ACTION LastComp_active:
wButtonColor:=16#FF00FFFF;

sStateDescription	:=	'Finish';
sStateInstructions	:= 	'LastComponentMixed';

bDisableAmount	:=FALSE;
bDisableName	:=FALSE;
bDisableTime	:=FALSE;
END_ACTION

ACTION LastComp_exit:
VisuElems.CurrentVisu:= 'StartVisu';
stTriblender.bDisolvingDone:=TRUE;
END_ACTION

ACTION MixComponent_active:
sStateDescription	:=	'Component Inside';
sStateInstructions	:= 	'Insert component in
 the specified amount';
END_ACTION

ACTION MixComponent_entry:
bContinue:=FALSE;

bDisableAmount	:=FALSE;
bDisableName	:=FALSE;
bDisableTime	:=FALSE;

wButtonColor:=16#FFFF0000;
IF iCurrentMixingComponent<g_Prod.cMaxCompInProduct-1 THEN
	stTriblender.bLastComponent:=NOT arrComponents[iCurrentMixingComponent+1].bComponentEnable;
END_IF
stTriblender.sComponenetAmount:=TO_STRING(arrComponents[iCurrentMixingComponent].rCompActWeight);
stTriblender.sComponenetName:=arrComponents[iCurrentMixingComponent].sDescription;
stTriblender.tComponenetMixingTime:=TO_TIME(arrComponents[iCurrentMixingComponent].iMixingTime*1000);
fb_TriBlenderPump.m_Run(RPM:=arrComponents[iCurrentMixingComponent].rRpmTarget);
END_ACTION

ACTION MixDoneWaitAnother_active:
sStateDescription	:='Triblender valve Opened';
sStateInstructions	:= 'Mix Component done,
 open triblender valve';
END_ACTION

ACTION MixDoneWaitAnother_entry:
bContinue:=FALSE;

bDisableAmount:=TRUE;
bDisableName:=TRUE;
bDisableTime:=TRUE;
bDisableButton:=FALSE;
VisuElems.CurrentVisu:= 'StartVisu';



wButtonColor:=16#FF00FF00;
END_ACTION

ACTION OpenValve_entry:
bContinue:=FALSE;

bDisableAmount:=TRUE;
bDisableName:=TRUE;
bDisableTime:=TRUE;
bDisableButton:=FALSE;

tonStageCirculation(IN:=FALSE);


sStateDescription	:='Triblender valve Opened';
sStateInstructions	:= 'Open triblender valve';

wButtonColor:=16#FF00FF00;
END_ACTION

TRANSITION trans_RpmInTarget:
fb_TriBlenderPump.nRPM< arrComponents[i].rRpmTarget+10 and fb_TriBlenderPump.nRPM> arrComponents[i].rRpmTarget-10
END_TRANSITION

TRANSITION transCircDone:
tonStageCirculation.Q and stTriblender.rMaxAllowedPressure> stTriblender.rPressure and stTriblender.rMinAllowedFlow< stTriblender.rFlow
END_TRANSITION

ACTION WaitForDone_active:
tonStageCirculation(IN:= TRUE,PT:=stTriblender.tComponenetMixingTime);
iCirculationTimeLeft:= TO_UINT(tonStageCirculation.PT - tonStageCirculation.ET)/1000;
bDisableButton:=TRUE;
END_ACTION

ACTION WaitForDone_entry:
wButtonColor:=16#FF0000FF;

sStateDescription	:=	'Waiting';
sStateInstructions	:= 	'Wait for mixing done';
bContinue:=FALSE;

bDisableAmount	:=FALSE;
bDisableName	:=FALSE;
bDisableTime	:=FALSE;


tonStageCirculation(IN:= FALSE);
END_ACTION

ACTION WaitForDone_exit:
stTriblender.bComponenetMixDone:=TRUE;
wButtonColor:=16#FF00FF00;

bDisableAmount	:=TRUE;
bDisableName	:=TRUE;
bDisableTime	:=TRUE;


tonStageCirculation(IN:= FALSE);
END_ACTION

ACTION WaitForStartPump_active:
sStateDescription	:='Start Water Circulation';
sStateInstructions	:= 'Start water circulation, check for leaks';
iCurrentMixingComponent:=0;
bContinue:=FALSE;
FOR i:= 0 TO g_Prod.cMaxCompInProduct-1 DO
	IF arrComponents[i].bIsWater THEN
		fb_TriBlenderPump.m_Run(RPM:=arrComponents[i].rRpmTarget);
	END_IF
END_FOR

wButtonColor:=16#FFFF0000;
END_ACTION

ACTION WaitForStartPump_entry:

stTriblender.bStartDisolving:=FALSE;
END_ACTION

ACTION WaterCirculation_active:
tonStageCirculation(IN:= stTriblender.bPumpOnFdbk,PT:=stTriblender.tWaterCirculationTimeout);
iCirculationTimeLeft:= TO_UINT(tonStageCirculation.PT - tonStageCirculation.ET)/1000;

bDisableButton:=TRUE;

sStateDescription	:='Wait for pressure and flow';
sStateInstructions	:= 'Water circulation in progress,
 check for leaks';
END_ACTION

ACTION WaterCirculation_entry:
bContinue:=FALSE;


bDisableAmount:=TRUE;
bDisableName:=TRUE;
bDisableTime:=FALSE;

tonStageCirculation(IN:=FALSE);
END_ACTION

ACTION WaterCirculation_exit:
tonStageCirculation(IN:=FALSE);
END_ACTION

END_PROGRAM

// ---- 03 Project/23 CIP/FB_Fill_Water.TcPOU
FUNCTION_BLOCK FB_Fill_Water EXTENDS FB_SFC_Cycle
VAR_INPUT
	valve : E_Pis_Name;;
	reqLevel: REAL;
	actLevel: REAL;
	
	fillCondition: BOOL;


END_VAR
VAR_OUTPUT
END_VAR
VAR
	fbHysteresis: FB_Hysteresis_REAL;
	stValve: REFERENCE TO ST_Piston;

END_VAR

stValve REF= stPis[valve];
IF NOT __ISVALIDREF(stValve) THEN;
	RETURN;
END_IF

fbHysteresis(
	fIn:= , 
	fHigh:= reqLevel, 
	fLow:= reqLevel-50.0, 
	iDigitsAfterDot:= , 
	bOut=> );

IF stValve.st_Open 
AND (NOT fbHysteresis.bOut
OR NOT fillCondition)
THEN;
	stValve.req_Close:=TRUE;
	
ELSIF stValve.st_Close 
AND fbHysteresis.bOut
THEN;
	stValve.req_Open:=TRUE;
END_IF

END_FUNCTION_BLOCK

// ---- 00 Library/01 Piston/TextList_Piston_Recipe_State.TcTLO
TEXTLIST TextList_Piston_Recipe_State
  0 = ' '
  1 = 'Open'
  2 = 'Close'
   = ''
END_TEXTLIST

// ---- 00 Library/01 Piston/TextList_Piston_Recipe_State_CloseOpen.TcTLO
TEXTLIST TextList_Piston_Recipe_State_CloseOpen
  0 = ' '
  1 = 'Close'
  2 = 'Open'
   = ''
END_TEXTLIST

// ---- 00 Library/01 Piston/TextList_Piston_Recipe_State_DownUp.TcTLO
TEXTLIST TextList_Piston_Recipe_State_DownUp
  0 = ' '
  1 = 'Down'
  2 = 'Up'
   = ''
END_TEXTLIST

// ---- 00 Library/01 Piston/TextList_Piston_Recipe_State_InOut.TcTLO
TEXTLIST TextList_Piston_Recipe_State_InOut
  0 = ' '
  1 = 'In'
  2 = 'Out'
   = ''
END_TEXTLIST

// ---- 00 Library/01 Piston/TextList_Piston_Recipe_State_OnOff.TcTLO
TEXTLIST TextList_Piston_Recipe_State_OnOff
  0 = ' '
  1 = 'On'
  2 = 'Off'
   = ''
END_TEXTLIST

// ---- 00 Library/01 Piston/TextList_Piston_Recipe_State_OpenClose.TcTLO
TEXTLIST TextList_Piston_Recipe_State_OpenClose
  0 = ' '
  1 = 'Open'
  2 = 'Close'
   = ''
END_TEXTLIST

// ---- 00 Library/01 Piston/TextList_Piston_Recipe_State_UpDown.TcTLO
TEXTLIST TextList_Piston_Recipe_State_UpDown
  0 = ' '
  1 = 'Up'
  2 = 'Down'
   = ''
END_TEXTLIST

// ---- 00 Library/01 Piston/VISU/vis_Piston_Control1.TcVIS
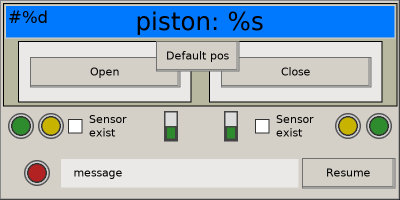
VISUALIZATION vis_Piston_Control1  // 400x200
VAR_IN_OUT
	stPis: ST_Piston;
END_VAR
    Rectangle (0,0 400x200)
    Rectangle (3,3 394x103), colour toggle: NOT stPis.b_Enable
    Rectangle (18,41 173x61), colour toggle: stPis.st_Open
    Rectangle (209,41 173x61), colour toggle: stPis.st_Close
    Button (30,57 150x30), "Open", colour toggle: stPis.req_Open, input disabled if: stPis.b_DeactivateMan OR NOT stPis.b_InterLock_Open
        toggle stPis.req_OpenMan
    Button (221,57 150x30), "Close", colour toggle: stPis.req_Close, input disabled if: stPis.b_DeactivateMan OR NOT stPis.b_InterLock_Close
        toggle stPis.req_CloseMan
    DipSwitch (156,111 30x30), tooltip "Open Sensor state", variable: stPis.sen_Open, invisible if: NOT stPis.sen_Open_Exist, behaviour: TOGGLE, style: Switch-DipSwitch-Green
    DipSwitch (216,111 30x30), tooltip "Close Sensor state", variable: stPis.sen_Close, invisible if: NOT stPis.sen_Close_Exist, behaviour: TOGGLE, style: Switch-DipSwitch-Green
    Checkbox (66,108 99x36), "Sensor exist", variable: stPis.sen_Open_Exist
    Checkbox (253,108 99x36), "Sensor exist", variable: stPis.sen_Close_Exist
    Lamp1 (6,111 30x30), tooltip "Open sensor", variable: stPis.sen_Open, invisible if: NOT stPis.sen_Open_Exist, style: Lamp-Lamp1-Green
    Lamp1 (333,111 30x30), tooltip "Close valve", variable: stPis.valve_Close, style: Lamp-Lamp1-Yellow
    Lamp1 (22,158 30x30), tooltip "Error", variable: stPis.b_Error, style: Lamp-Lamp1-Red
    Textfield (60,158 239x30), "message"
    Button (302,158 93x30), "Resume", colour toggle: stPis.b_Error
        toggle stPis.b_Resume
    Button (156,41 83x30), "Default pos", colour toggle: stPis.req_DefaultPos, input disabled if: stPis.b_DeactivateMan
        toggle stPis.req_DefaultPos
    Textfield (5,5 390x33), "piston: %s", text variable: stPis.sName
    Textfield (5,7 42x21), "#%d", text variable: stPis.iPisNum
    Lamp1 (36,111 30x30), tooltip "Open valve", variable: stPis.valve_Open, style: Lamp-Lamp1-Yellow
    Lamp1 (364,111 30x30), tooltip "Close sensor", variable: stPis.sen_Close, invisible if: NOT stPis.sen_Close_Exist, style: Lamp-Lamp1-Green
END_VISUALIZATION

// ---- 00 Library/01 Piston/VISU/vis_Piston_Control1_Compact.TcVIS
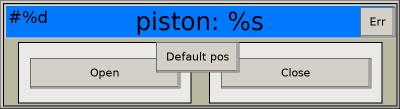
VISUALIZATION vis_Piston_Control1_Compact  // 400x109
VAR_IN_OUT
	stPis: ST_Piston;
END_VAR
    Rectangle (0,0 400x109)
    Rectangle (3,3 394x103), colour toggle: NOT stPis.b_Enable
    Rectangle (18,42 173x61), colour toggle: stPis.st_Open
    Rectangle (209,42 173x61), colour toggle: stPis.st_Close
    Button (30,58 150x30), "Open", colour toggle: stPis.req_Open, input disabled if: stPis.b_DeactivateMan OR NOT stPis.b_InterLock_Open
        toggle stPis.req_OpenMan
    Button (221,58 150x30), "Close", colour toggle: stPis.req_Close, input disabled if: stPis.b_DeactivateMan OR NOT stPis.b_InterLock_Close
        toggle stPis.req_CloseMan
    Button (156,42 83x30), "Default pos", colour toggle: stPis.req_DefaultPos, input disabled if: stPis.b_DeactivateMan
        toggle stPis.req_DefaultPos
    Textfield (5,5 390x33), "piston: %s", text variable: stPis.sName
    Textfield (5,7 42x21), "#%d", text variable: stPis.iPisNum
    Button (360,7 35x30), "Err", colour toggle: stPis.b_Error
        toggle stPis.b_Resume
END_VISUALIZATION

// ---- 00 Library/01 Piston/VISU/vis_Piston_Control2_CloseOpen.TcVIS
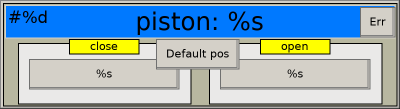
VISUALIZATION vis_Piston_Control2_CloseOpen  // 400x109
VAR_IN_OUT
	stPis			: ST_Piston;
END_VAR
VAR_INPUT
	sLable_Open		: STRING:='lable open';
	sLable_Close	: STRING:='lable close';
END_VAR
    Rectangle (0,0 400x109)
    Rectangle (3,3 394x103), colour toggle: NOT stPis.b_Enable
    Rectangle (209,43 173x61), colour toggle: stPis.st_Open
    Button (220,59 150x30), "%s", text variable: sLable_Open, colour toggle: stPis.req_Open, input disabled if: stPis.b_DeactivateMan OR NOT stPis.b_InterLock_Open
        toggle stPis.req_OpenMan
    RoundedRectangle (260,39 70x15), "open"
    Rectangle (18,43 173x61), colour toggle: stPis.st_Close
    Button (29,59 150x30), "%s", text variable: sLable_Close, colour toggle: stPis.req_Close, input disabled if: stPis.b_DeactivateMan OR NOT stPis.b_InterLock_Close
        toggle stPis.req_CloseMan
    RoundedRectangle (69,39 70x15), "close"
    Button (156,39 83x30), "Default pos", colour toggle: stPis.req_DefaultPos, input disabled if: stPis.b_DeactivateMan
        toggle stPis.req_DefaultPos
    Textfield (5,5 390x33), "piston: %s", text variable: stPis.description
    Textfield (5,7 42x21), "#%d", text variable: stPis.iPisNum
    Button (360,7 35x30), "Err", colour toggle: stPis.b_Error
        toggle stPis.b_Resume
END_VISUALIZATION

// ---- 00 Library/01 Piston/VISU/vis_Piston_Control2_OpenClose.TcVIS
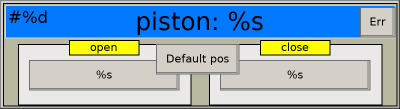
VISUALIZATION vis_Piston_Control2_OpenClose  // 400x109
VAR_IN_OUT
	stPis			: ST_Piston;
END_VAR
VAR_INPUT
	sLable_Open		: STRING:='lable open';
	sLable_Close	: STRING:='lable close';
END_VAR
    Rectangle (0,0 400x109)
    Rectangle (3,3 394x103), colour toggle: NOT stPis.b_Enable
    Rectangle (18,44 173x61), colour toggle: stPis.st_Open
    Rectangle (209,44 173x61), colour toggle: stPis.st_Close
    Button (29,60 150x30), "%s", text variable: sLable_Open, colour toggle: stPis.req_Open, input disabled if: stPis.b_DeactivateMan OR NOT stPis.b_InterLock_Open
        toggle stPis.req_OpenMan
    Button (220,60 150x30), "%s", text variable: sLable_Close, colour toggle: stPis.req_Close, input disabled if: stPis.b_DeactivateMan OR NOT stPis.b_InterLock_Close
        toggle stPis.req_CloseMan
    Button (156,44 83x30), "Default pos", colour toggle: stPis.req_DefaultPos, input disabled if: stPis.b_DeactivateMan
        toggle stPis.req_DefaultPos
    RoundedRectangle (69,40 70x15), "open"
    RoundedRectangle (260,40 70x15), "close"
    Textfield (5,5 390x33), "piston: %s", text variable: stPis.description
    Textfield (5,7 42x21), "#%d", text variable: stPis.iPisNum
    Button (360,7 35x30), "Err", colour toggle: stPis.b_Error
        toggle stPis.b_Resume
END_VISUALIZATION

// ---- 00 Library/01 Piston/VISU/vis_Piston_Select.TcVIS
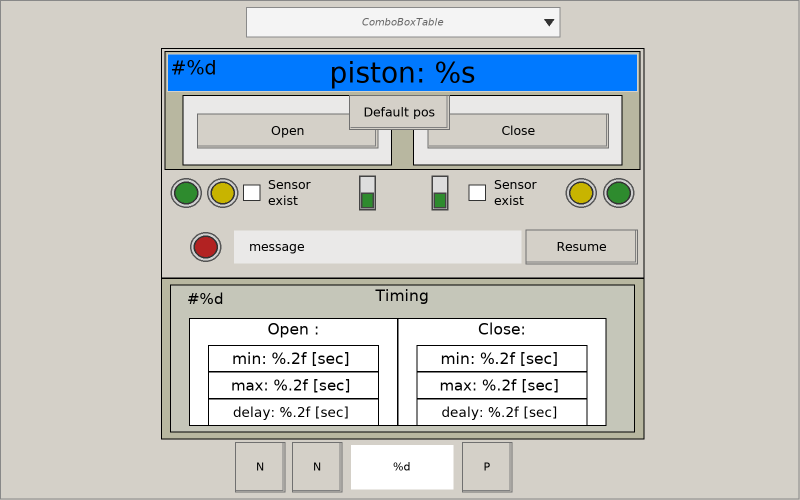
VISUALIZATION vis_Piston_Select  // 800x500
    Frame (161,48 483x230)
        shows vis_Piston_Control1(stPis := stPis[iPis_sel])
    Frame (161,278 483x161)
        shows vis_Piston_Times(stPis := stPis[iPis_sel])
    Button (292,442 50x50), "N"
        tap prg_Piston.bPis_Next_N
    Button (462,442 50x50), "P"
        tap prg_Piston.bPis_Next_P
    Textfield (350,444 104x46), "%d", text variable: iPis_sel
    ComboBoxTable (246,7 314x30), variable: iPis_sel, data array: g_Piston.arPisName
        p3854506369: g_Piston.arPisName[INDEX].Num
        p1892666644: g_Piston.arPisName[INDEX].Description
    Button (235,442 50x50), "N"
        tap prg_Piston.bPis_Next_N
END_VISUALIZATION

// ---- 00 Library/01 Piston/VISU/vis_Piston_Select_1.TcVIS
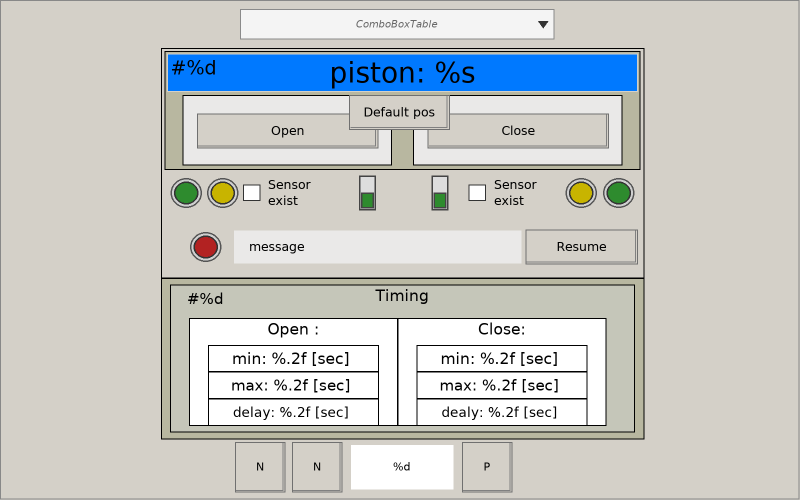
VISUALIZATION vis_Piston_Select_1  // 800x500
    Frame (161,48 483x230)
        shows vis_Piston_Control1(stPis := stPis[iPis_sel])
    Frame (161,278 483x161)
        shows vis_Piston_Times(stPis := stPis[iPis_sel])
    Button (292,442 50x50), "N"
        tap prg_Piston.bPis_Next_N
    Button (462,442 50x50), "P"
        tap prg_Piston.bPis_Next_P
    Textfield (350,444 104x46), "%d", text variable: iPis_sel
    ComboBoxTable (240,9 314x30), variable: iPis_sel, data array: arPisName
        p1128707560: C_MAX_Pistons_Exist
        p3854506369: arPisName[INDEX].Num
        p1892666644: arPisName[INDEX].Description
    Button (235,442 50x50), "N"
        tap prg_Piston.bPis_Next_N
END_VISUALIZATION

// ---- 00 Library/01 Piston/VISU/vis_Piston_Setting_Table.TcVIS
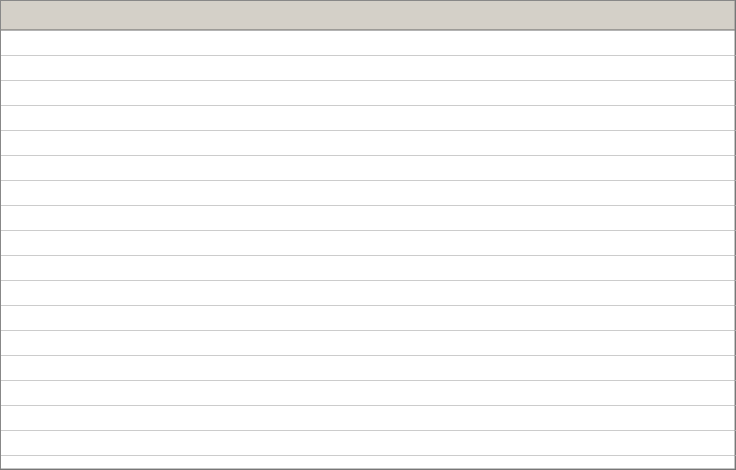
VISUALIZATION vis_Piston_Setting_Table  // 736x470
    Table (0,0 736x470), data array: stPisSetting
        p3854506369: stPisSetting[INDEX].t_minOpen
        p1892666644: stPisSetting[INDEX].t_minClose
        p338671338: stPisSetting[INDEX].t_maxOpen
        p2170511999: stPisSetting[INDEX].t_maxClose
        p3723444502: stPisSetting[INDEX].t_DelayOpen
        p1218418051: stPisSetting[INDEX].t_DelayClose
        p746581629: stPisSetting[INDEX].sen_Open_Exist
        p3104783080: stPisSetting[INDEX].sen_Close_Exist
END_VISUALIZATION

// ---- 00 Library/01 Piston/VISU/vis_Piston_Times.TcVIS
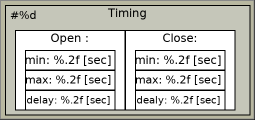
VISUALIZATION vis_Piston_Times  // 255x120
VAR_IN_OUT
	stPis: ST_Piston;
END_VAR
    Rectangle (0,0 255x120)
    Rectangle (5,5 245x110), "Timing"
    Rectangle (15,30 110x80), "Open :"
    Rectangle (125,30 110x80), "Close:"
    Rectangle (135,50 90x20), "min: %.2f [sec]", text variable: stPis.t_minClose
        OnMouseDown: write the text variable via Edit, min 0
    Rectangle (135,70 90x20), "max: %.2f [sec]", text variable: stPis.t_maxClose
        OnMouseDown: write the text variable via Edit, min 0
    Rectangle (25,70 90x20), "max: %.2f [sec]", text variable: stPis.t_maxOpen
        OnMouseDown: write the text variable via Edit, min 0
    Rectangle (25,50 90x20), "min: %.2f [sec]", text variable: stPis.t_minOpen
        OnMouseDown: write the text variable via Edit, min 0
    Rectangle (25,90 90x20), "delay: %.2f [sec]", text variable: stPis.t_DelayOpen
        OnMouseDown: write the text variable via Edit, min 0
    Rectangle (135,90 90x20), "dealy: %.2f [sec]", text variable: stPis.t_DelayClose
        OnMouseDown: write the text variable via Edit, min 0
    Textfield (4,5 39x21), "#%d", text variable: stPis.iPisNum
END_VISUALIZATION

// ---- 00 Library/03 SFC/vis_Cycle_Control.TcVIS
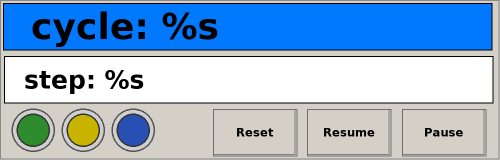
VISUALIZATION vis_Cycle_Control  // 500x160
VAR_IN_OUT
	fb: FB_SFC_Cycle;
END_VAR
VAR_INPUT
	sName: STRING:='Cycle name';
END_VAR
    Lamp1 (8,105 50x50), tooltip "Ready", variable: fb.bReady, style: Lamp-Lamp1-Green
    Lamp1 (108,105 50x50), tooltip "Done", variable: fb.bDone, style: Lamp-Lamp1-Blue
    Lamp1 (58,105 50x50), tooltip "Run", variable: fb.bRun, style: Lamp-Lamp1-Yellow
    RoundedRectangle (3,3 489x47), "cycle: %s", tooltip "POU name: %s", text variable: sName
        p4168582468: fb.refSFC.SFCErrorPOU
    RoundedRectangle (4,56 489x47), "step: %s", text variable: fb.refSFC.SFCCurrentStep, colour toggle: fb.ErrorSFC
    Button (213,109 84x47), "Reset"
        tap fb.bInit
    Button (307,109 84x47), "Resume", colour toggle: fb.ErrorSFC
        toggle fb.refSFC.SFCQuitError
    Button (402,109 84x47), "Pause", colour toggle: fb.refSFC.SFCPause
        toggle fb.refSFC.SFCPause
END_VISUALIZATION

// ---- 00 Library/03 SFC/vis_Cycle_Control_1.TcVIS
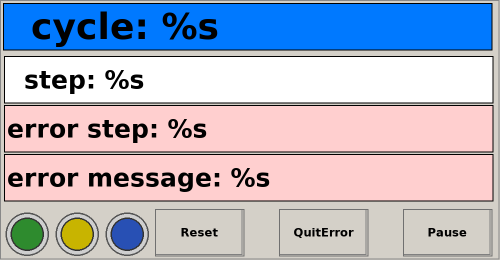
VISUALIZATION vis_Cycle_Control_1  // 500x260
VAR_IN_OUT
	fb: FB_SFC_Cycle;
END_VAR
VAR_INPUT
	sName: STRING:='Cycle name';
END_VAR
    Lamp1 (2,209 50x50), tooltip "Ready", variable: fb.bReady, style: Lamp-Lamp1-Green
    Lamp1 (102,209 50x50), tooltip "Done", variable: fb.bDone, style: Lamp-Lamp1-Blue
    Lamp1 (52,209 50x50), tooltip "Run", variable: fb.bRun, style: Lamp-Lamp1-Yellow
    RoundedRectangle (3,3 489x47), "cycle: %s", tooltip "POU name: %s", text variable: sName
        p4168582468: fb.refSFC.SFCErrorPOU
    RoundedRectangle (4,56 489x47), "step: %s", text variable: fb.refSFC.SFCCurrentStep, colour toggle: fb.ErrorSFC
    Button (155,209 89x47), "Reset"
        tap fb.bInit
    Button (403,209 89x47), "Pause", colour toggle: fb.refSFC.SFCPause
        toggle fb.refSFC.SFCPause
    Button (279,209 89x47), "QuitError", colour toggle: fb.ErrorSFC
        toggle fb.refSFC.SFCQuitError
    RoundedRectangle (4,105 489x47), "error step: %s", text variable: fb.sLastStepBefore_Error, colour toggle: fb.ErrorSFC
    RoundedRectangle (4,154 489x47), "error message: %s", text variable: fb.sError_Message, colour toggle: fb.ErrorSFC
END_VISUALIZATION

// ---- 00 Library/03 SFC/vis_Cycle_Panel.TcVIS
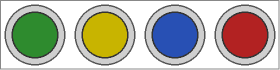
VISUALIZATION vis_Cycle_Panel  // 280x70
VAR_IN_OUT
	fb: FB_SFC_Cycle;
END_VAR
    Lamp1 (0,0 70x70), tooltip "Ready", variable: fb.bReady, style: Lamp-Lamp1-Green
    Lamp1 (70,0 70x70), tooltip "Done", variable: fb.bDone, style: Lamp-Lamp1-Yellow
    Lamp1 (140,0 70x70), tooltip "ToBe Done", variable: fb.bToBe_Done, style: Lamp-Lamp1-Blue
    Lamp1 (210,0 70x70), tooltip "Run", variable: fb.bRun, style: Lamp-Lamp1-Red
END_VISUALIZATION

// ---- 00 Library/04 Recipe/FB_Recipe_Vizu.TcVIS
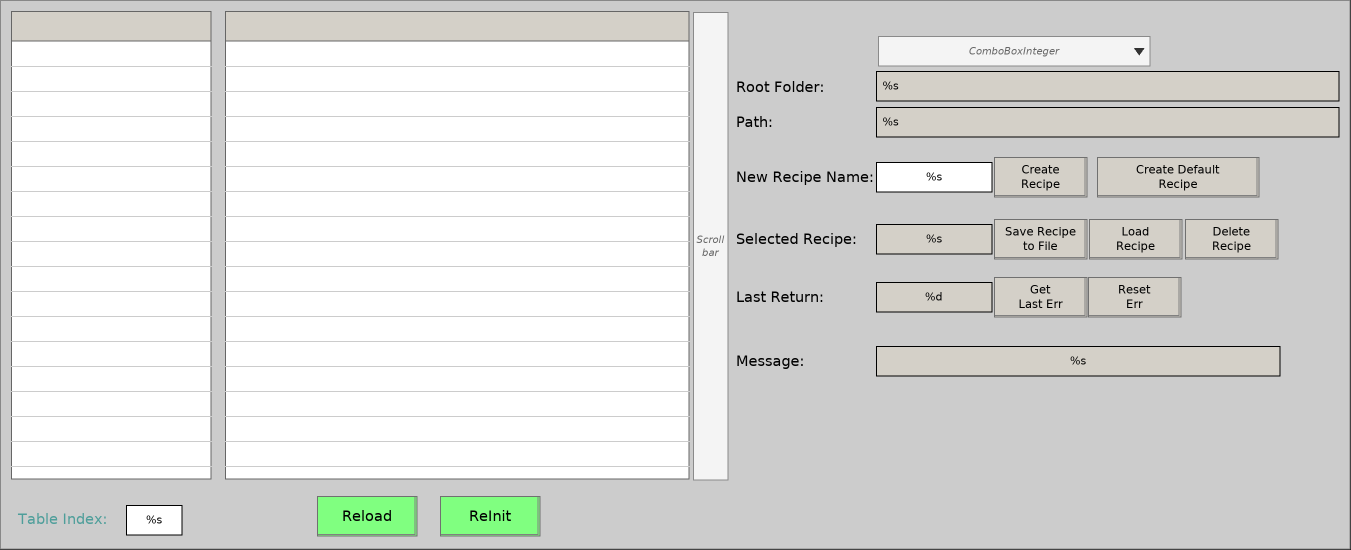
VISUALIZATION FB_Recipe_Vizu  // 1351x550
VAR_IN_OUT
	fb_Recipe		:FB_Recipe;
END_VAR
    Rectangle (0,0 1351x550)
    Table (11,11 200x468), data array: fb_Recipe.pstRecipe^.arrRecipeNames
        p1137915858: fb_Recipe.pstRecipe^.iRecipeIndex
        p1822360349: fb_Recipe.pstRecipe^.bValidSelected
        p3854506369: fb_Recipe.pstRecipe^.arrRecipeNames[INDEX]
        p2232123230: Recipe Names
    Rectangle (126,505 56x30), "%s", text variable: fb_Recipe.pstRecipe^.iRecipeIndex
    Label (15,504 108x30), "Table Index:"
    Button (317,496 100x40), "Reload"
        toggle fb_Recipe.pstRecipe^.bReloadRecipes
    Table (225,11 464x468), data array: fb_Recipe.pstRecipe^.arrVariableDisp
        p3854506369: fb_Recipe.pstRecipe^.arrVariableDisp[0,INDEX]
        p2232123230: No
        p1892666644: fb_Recipe.pstRecipe^.arrVariableDisp[1,INDEX]
        p511219082: Variable Name
        p338671338: fb_Recipe.pstRecipe^.arrVariableDisp[2,INDEX]
        p1755163831: Variable Value
    Scrollbar (693,12 35x468)
        p1057716461: fb_Recipe.pstRecipe^.iDispSel
    Button (1185,219 93x40), "Delete Recipe"
        toggle fb_Recipe.pstRecipe^.bDeleteRecipe
    Label (733,162 141x30), "New Recipe Name:"
    Label (733,224 141x30), "Selected Recipe:"
    Label (733,282 141x30), "Last Return:"
    Rectangle (876,162 116x30), "%s", text variable: fb_Recipe.pstRecipe^.sNewRecipeName
        OnMouseClick: write the text variable via Edit
    Rectangle (876,224 116x30), "%s", text variable: fb_Recipe.pstRecipe^.sSelectedReceipe
    Rectangle (876,282 116x30), "%d", text variable: fb_Recipe.LastReturn, colour toggle: fb_Recipe.LastReturn<>0
    Button (994,157 93x40), "Create Recipe"
        toggle fb_Recipe.pstRecipe^.bCreateRecipe
    Button (994,219 93x40), "Save Recipe to File"
        toggle fb_Recipe.pstRecipe^.bSaveFileCmd
    Button (994,277 93x40), "Get Last Err"
        toggle fb_Recipe.pstRecipe^.bGetLastError
    Button (1089,219 93x40), "Load Recipe"
        toggle fb_Recipe.pstRecipe^.bWriteToPLC_Cmd
    Button (1088,277 93x40), "Reset Err"
        toggle fb_Recipe.pstRecipe^.bResetLastError
    Label (733,107 141x30), "Path:"
    Rectangle (876,107 463x30), "%s", text variable: fb_Recipe.sRecipesStoragePath
    Button (440,496 100x40), "ReInit"
        toggle fb_Recipe.pstRecipe^.bReInit
    Label (733,346 141x30), "Message:"
    Rectangle (876,346 404x30), "%s", text variable: fb_Recipe.sMessage
    Button (1097,157 162x40), "Create Default Recipe"
        toggle fb_Recipe.pstRecipe^.bCreateRecipe
        OnMouseClick: execute { fb_Recipe.pstRecipe^.sNewRecipeName:='Default'; }
    ComboBoxInteger (878,36 272x30), variable: GVL_Recipe.eRecipeRootFolder, text list: 'TextList_RecipeRootFolder'
    Rectangle (876,71 463x30), "%s", text variable: GVL_Recipe.ar_RecipesStoragePath_Root[GVL_Recipe.eRecipeRootFolder]
        OnMouseClick: write the text variable via Edit
    Label (733,72 141x30), "Root Folder:"
END_VISUALIZATION

// ---- 00 Library/04 Recipe/OLD/vis_RecipeControl_v01.TcVIS
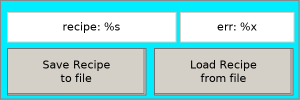
VISUALIZATION vis_RecipeControl_v01  // 300x100
VAR_INPUT
	Definition: STRING;
END_VAR
VAR
	RecipeName: STRING:='name';
END_VAR
    Button (7,48 139x47), "Save Recipe to file"
        OnMouseClick: ExecuteCommand ExecuteCommand=ExecuteCommand=[Command=CreateRecipe, Value=Definition, Value2=RecipeName, Command=SaveRecipeAs, Value=Definition, Value2=RecipeName]
    Button (154,48 139x47), "Load Recipe from file"
        OnMouseClick: ExecuteCommand ExecuteCommand=ExecuteCommand=[Command=LoadRecipeFrom, Value=Definition, Value2=RecipeName]
    Textfield (7,12 169x30), "recipe: %s", text variable: Definition
    Textfield (180,12 114x30), "err: %x", text variable: prg_RecipeManager.LastError, colour toggle: prg_RecipeManager.LastError<>0
        toggle prg_RecipeManager.bResetError
END_VISUALIZATION

// ---- 00 Library/04 Recipe/OLD/vis_RecipeTest.TcVIS
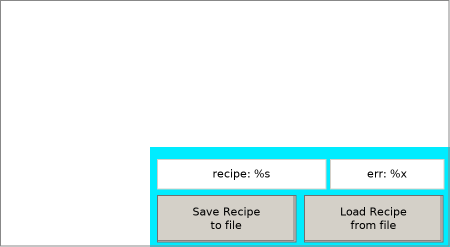
VISUALIZATION vis_RecipeTest  // 450x247
    Frame (150,147 300x100)
        shows vis_RecipeControl_v01(Definition := 'R_Open1')
END_VISUALIZATION

// ---- 00 Library/04 Recipe/TextList_RecipeRootFolder.TcTLO
TEXTLIST TextList_RecipeRootFolder
  0 = 'PLC'
  1 = 'Develop 1'
  2 = 'Develop 2'
  3 = 'Develop 3'
  4 = 'Develop 4'
   = ''
END_TEXTLIST

// ---- 00 Library/05 Safety/Vis_ES_PB.TcVIS
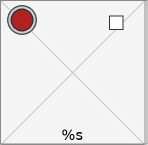
VISUALIZATION Vis_ES_PB  // 148x145
VAR_IN_OUT
	stPB: ST_ES_PB;

END_VAR
VAR_INPUT
	Lable: STRING;

END_VAR
    Image (0,0 145x145), "%s", text variable: Lable, image: ImagePool.EStop_OK2
        p84334746: stPB.stBitMap
    Checkbox (107,3 41x39), tooltip "ByPass", variable: stPB.ByPass, input disabled if: prg_User.actUser<4
    Lamp1 (5,3 34x34), tooltip "Memo PB State", variable: stPB.Memo, style: Lamp-Lamp1-Red
END_VISUALIZATION

// ---- 00 Library/06-Visu/Sensor.TcVIS
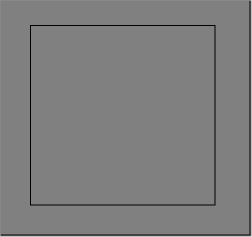
VISUALIZATION Sensor  // 252x237
VAR_INPUT
	{attribute 'parameterstringof' := 'm_Input_Sen_Addr'}
	m_Input_Sen_Addr_Str : STRING;
END_VAR
VAR_INPUT
	m_Input_Sen_Addr : Bool;
END_VAR
    Rectangle (0,0 250x235)
    RoundedRectangle (30,25 185x180), tooltip "%s", colour toggle: (m_Input_Sen_Addr) <> 0
        p4168582468: m_Input_Sen_Addr_Str
END_VISUALIZATION

// ---- 00 Library/07 Errors/vis_Device_Error.TcVIS
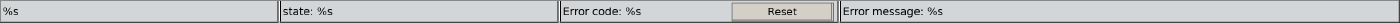
VISUALIZATION vis_Device_Error  // 1500x25
VAR_IN_OUT
	fb_comm_dev: fb_common_device;
END_VAR
    Rectangle (900,0 600x25), "Error message: %s", text variable: fb_comm_dev.common_events.device_error.error_string, colour toggle: fb_comm_dev.common_events.device_error.error_code<>''
        OnMouseUp: execute { GVL.Errors:=(0); }
    Rectangle (600,0 298x25), "Error code: %s", text variable: fb_comm_dev.common_events.device_error.error_code, colour toggle: fb_comm_dev.common_events.device_error.error_code<>''
        OnMouseUp: execute { GVL.Errors:=(0); }
    Button (784,3 109x20), "Reset"
        toggle fb_comm_dev.common_actions.reset
    Rectangle (0,0 298x25), "%s", tooltip "Device Name", text variable: fb_comm_dev.Name, colour toggle: fb_comm_dev.common_events.device_error.error_code<>''
        OnMouseUp: execute { GVL.Errors:=(0); }
    Rectangle (300,0 298x25), "state: %s", tooltip "Device State", text variable: fb_comm_dev.device_status, colour toggle: fb_comm_dev.common_events.device_error.error_code<>''
        OnMouseUp: execute { GVL.Errors:=(0); }
END_VISUALIZATION

// ---- 00 Library/07-Mode/Visu/Mode_Select.TcVIS
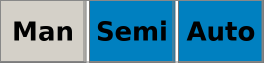
VISUALIZATION Mode_Select  // 264x63
VAR_IN_OUT
	stMode: ST_Mode;
END_VAR
    Button (0,0 86x63), "Man", colour toggle: stModeMain.iActMode=eManualMode
        OnMouseDown: execute {
            stModeMain.bSetManual:=TRUE;
            stMode.bSetSemi:=FALSE;
            stMode.bSetAuto:=FALSE;
        }
    Button (89,0 86x63), "Semi", colour toggle: stModeMain.iActMode=eSemiAutoMode
        OnMouseDown: execute {
            stModeMain.bSetManual:=FALSE;
            stMode.bSetSemi:=TRUE;
            stMode.bSetAuto:=FALSE;
        }
    Button (178,0 86x63), "Auto", colour toggle: stModeMain.iActMode=eAutoMode
        OnMouseDown: execute {
            stModeMain.bSetManual:=FALSE;
            stMode.bSetSemi:=FALSE;
            stMode.bSetAuto:=TRUE;
        }
END_VISUALIZATION

// ---- 00 Library/07-Mode/Visu/Mode_Select_1.TcVIS
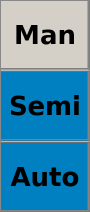
VISUALIZATION Mode_Select_1  // 90x212
VAR_IN_OUT
	stMode: ST_Mode;
END_VAR
    Button (0,0 90x70), "Man", colour toggle: stModeMain.iActMode=eManualMode, input disabled if: NOT GVL.MainMachine.bReadyToManualModeSelect
        OnMouseDown: execute {
            stModeMain.bSetManual:=TRUE;
            stMode.bSetSemi:=FALSE;
            stMode.bSetAuto:=FALSE;
        }
    Button (0,71 90x70), "Semi", colour toggle: stModeMain.iActMode=eSemiAutoMode, input disabled if: stModeMain.iActMode<>E_WorkingMode.eManualMode
        OnMouseDown: execute {
            stModeMain.bSetManual:=FALSE;
            stMode.bSetSemi:=TRUE;
            stMode.bSetAuto:=FALSE;
        }
    Button (0,142 90x70), "Auto", colour toggle: stModeMain.iActMode=eAutoMode, input disabled if: stModeMain.iActMode<>E_WorkingMode.eManualMode
        OnMouseDown: execute {
            stModeMain.bSetManual:=FALSE;
            stMode.bSetSemi:=FALSE;
            stMode.bSetAuto:=TRUE;
        }
END_VISUALIZATION

// ---- 00 Library/07-Mode/Visu/OperationButtons.TcVIS
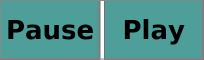
VISUALIZATION OperationButtons  // 204x60
VAR_IN_OUT
	stOperation	:ST_OperationButtons;
END_VAR
    Button (0,0 100x60), "Pause", tooltip "%s", colour toggle: stOperation.iActOperation=ePauseAll
        p4168582468: stOperation.sModeZone
        OnMouseClick: execute { stOperation.bSetPause:=TRUE; stOperation.iPauseHistory:=7; }
    Button (104,0 100x60), "Play", tooltip "%s", colour toggle: stOperation.iActOperation=ePlayAll
        p4168582468: stOperation.sModeZone
        OnMouseClick: execute { stOperation.bSetPlay:=TRUE; }
END_VISUALIZATION

// ---- 00 Library/07-Mode/Visu/OperationButtons_1.TcVIS
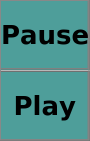
VISUALIZATION OperationButtons_1  // 90x141
VAR_IN_OUT
	stOperation	:ST_OperationButtons;
END_VAR
    Button (0,0 90x70), "Pause", colour toggle: stOperation.iActOperation=ePauseAll
        OnMouseClick: execute { stOperation.bSetPause:=TRUE; stOperation.iPauseHistory:=7; }
    Button (0,71 90x70), "Play", colour toggle: stOperation.iActOperation=ePlayAll
        OnMouseClick: execute { stOperation.bSetPlay:=TRUE; }
END_VISUALIZATION

// ---- 00 Library/07-Mode/Visu/OperationButton_Stop.TcVIS
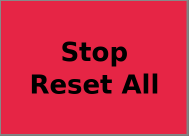
VISUALIZATION OperationButton_Stop  // 189x136
VAR_IN_OUT
	stOperation	:ST_OperationButtons;
END_VAR
    Button (0,0 189x136), "Stop Reset All", colour toggle: stOperation.bStopResetAll, pressed state: stOperation.bStopResetAll
        OnMouseClick: execute { stOperation.bStopResetAll:=TRUE; stOperation.iPauseHistory:=5; }
END_VISUALIZATION

// ---- 00 Library/07-Mode/Visu/Vis_PauseHistory.TcVIS
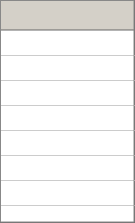
VISUALIZATION Vis_PauseHistory  // 135x223
VAR_IN_OUT
	fbOp: FB_Operation;
END_VAR
    Table (0,0 135x223), data array: fbOp.arPauseHistory
        p3854506369: fbOp.arPauseHistory[INDEX]
        p2232123230: Pause History
END_VISUALIZATION

// ---- 00 Library/10 Utils/DutyCycle/vis_FB_DutyCycle.TcVIS
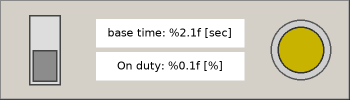
VISUALIZATION vis_FB_DutyCycle  // 350x100
VAR_IN_OUT
	fb: FB_DutyCycle;
END_VAR
    Rectangle (0,0 350x100)
    Lamp1 (266,15 70x70), variable: fb.bOut, style: Lamp-Lamp1-Yellow
    DipSwitch (10,15 70x70), variable: fb.bEnable, behaviour: TOGGLE, style: Switch-DipSwitch-Gray
    Textfield (95,18 150x30), "base time: %2.1f [sec]", text variable: fb.fBaseTime, input disabled if: prg_User.actUser<4
        OnMouseClick: write the text variable via Edit, min 0, max 60
    Textfield (95,51 150x30), "On duty: %0.1f [%]", text variable: fb.fOn_Duty
        OnMouseClick: write the text variable via Edit, min 0, max 100
END_VISUALIZATION

// ---- 00 Library/10 Utils/DutyCycle/vis_FB_DutyCycle_Master.TcVIS
